FUNCTION_BLOCK TableDriver (* Composite Function Block Type *)
  (* Standard: 61499-2 *)
  (* Version 0.0, 7/2/2026, template *)
  PACKAGE Main;
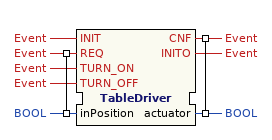
  EVENT_INPUT
    INIT; (* Initialization Request *)
    REQ WITH inPosition; (* Normal Execution Request *)
    TURN_ON;
    TURN_OFF;
  END_EVENT
  EVENT_OUTPUT
    CNF WITH actuator; (* Execution Confirmation *)
    INITO; (* Initialization Confirm *)
  END_EVENT
  VAR_INPUT
    inPosition : BOOL; (* Input event qualifier *)
  END_VAR
  VAR_OUTPUT
    actuator : BOOL; (* Output event qualifier *)
  END_VAR
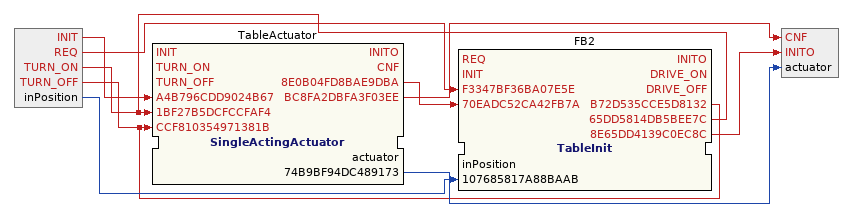
  FBS
    TableActuator : SingleActingActuator;
    FB2 : TableInit;
  END_FBS
  EVENT_CONNECTIONS
    REQ TO FB2.F3347BF36BA07E5E;
    INIT TO TableActuator.A4B796CDD9024B67;
    TURN_ON TO TableActuator.1BF27B5DCFCCFAF4;
    TURN_OFF TO TableActuator.CCF810354971381B;
    FB2.B72D535CCE5D8132 TO TableActuator.CCF810354971381B;
    FB2.65DD5814DB5BEE7C TO TableActuator.1BF27B5DCFCCFAF4;
    TableActuator.8E0B04FD8BAE9DBA TO FB2.70EADC52CA42FB7A;
    TableActuator.BC8FA2DBFA3F03EE TO CNF;
    FB2.8E65DD4139C0EC8C TO INITO;
  END_CONNECTIONS
  DATA_CONNECTIONS
    inPosition TO FB2.107685817A88BAAB;
    TableActuator.74B9BF94DC489173 TO actuator;
  END_CONNECTIONS
END_FUNCTION_BLOCK
